{attribute 'qualified_only'}
VAR_GLOBAL CONSTANT
    // Physical I/O interface is reserved; enable only after actual I/O mapping.
    ACTIVE_EXIO : BOOL := FALSE;
END_VAR

(* stored: Version 1.1.0.1, ProductVersion 3.1.4024.12
   GVL Config: Id {a7f3d0b1-8542-4197-8f4a-d81bdb596a28} *)
